(* Communikation structure from gefran to plc *)

TYPE ST_PLCTOGFX4IR_1 :
STRUCT
	nLocalSetPoint			:INT;
	nManualOutput			:WORD;
	wControllerStatus		:WORD;
END_STRUCT
END_TYPE

(* stored: Version 1.1.0.1, ProductVersion 3.1.4024.15
   DUT ST_PLCTOGFX4IR_1: Id {4197b7de-c932-4dec-a5c7-a139597785f1} *)
